// Mitsubishi GX Works2 project: 프로젝트1   PLC: Q03UDV

PROGRAM MAIN
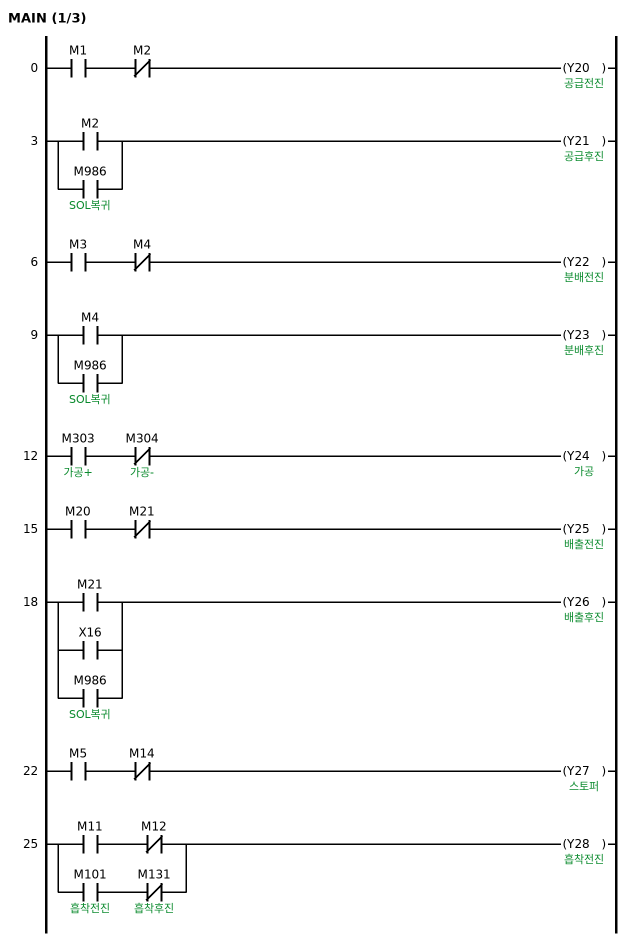
0     LD      M1
      ANI     M2
      OUT     Y20  ; 공급전진
3     LD      M2
      OR      M986  ; SOL복귀
      OUT     Y21  ; 공급후진
6     LD      M3
      ANI     M4
      OUT     Y22  ; 분배전진
9     LD      M4
      OR      M986  ; SOL복귀
      OUT     Y23  ; 분배후진
12    LD      M303  ; 가공+
      ANI     M304  ; 가공-
      OUT     Y24  ; 가공
15    LD      M20
      ANI     M21
      OUT     Y25  ; 배출전진
18    LD      M21
      OR      X16
      OR      M986  ; SOL복귀
      OUT     Y26  ; 배출후진
22    LD      M5
      ANI     M14
      OUT     Y27  ; 스토퍼
25    LD      M11
      ANI     M12
      LD      M101  ; 흡착전진
      ANI     M131  ; 흡착후진
      ORB
      OUT     Y28  ; 흡착전진
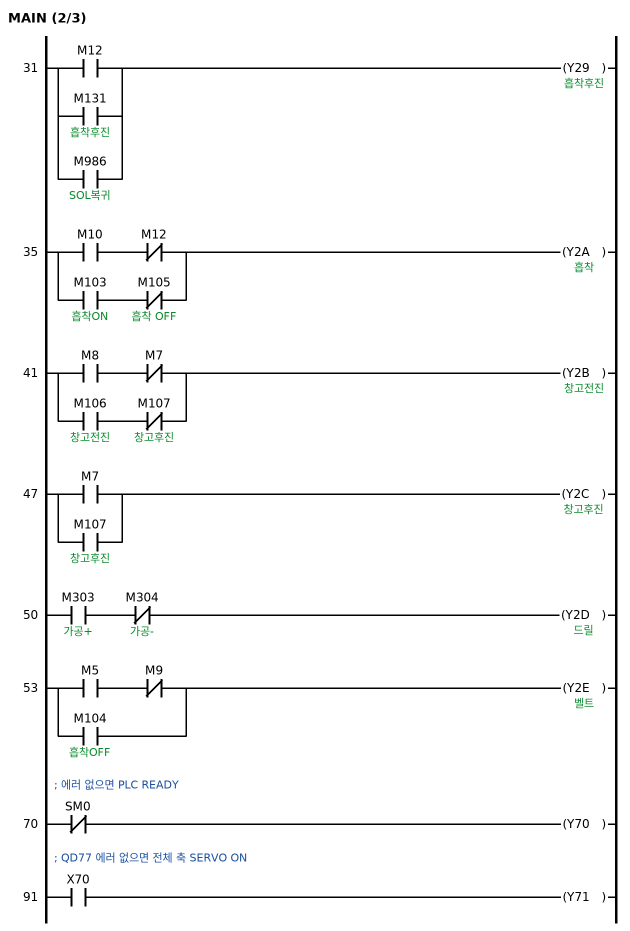
31    LD      M12
      OR      M131  ; 흡착후진
      OR      M986  ; SOL복귀
      OUT     Y29  ; 흡착후진
35    LD      M10
      ANI     M12
      LD      M103  ; 흡착ON
      ANI     M105  ; 흡착 OFF
      ORB
      OUT     Y2A  ; 흡착
41    LD      M8
      ANI     M7
      LD      M106  ; 창고전진
      ANI     M107  ; 창고후진
      ORB
      OUT     Y2B  ; 창고전진
47    LD      M7
      OR      M107  ; 창고후진
      OUT     Y2C  ; 창고후진
50    LD      M303  ; 가공+
      ANI     M304  ; 가공-
      OUT     Y2D  ; 드릴
53    LD      M5
      ANI     M9
      OR      M104  ; 흡착OFF
      OUT     Y2E  ; 벨트
; 에러 없으면 PLC READY
70    LDI     SM0
      OUT     Y70
; QD77 에러 없으면 전체 축 SERVO ON
91    LD      X70
      OUT     Y71
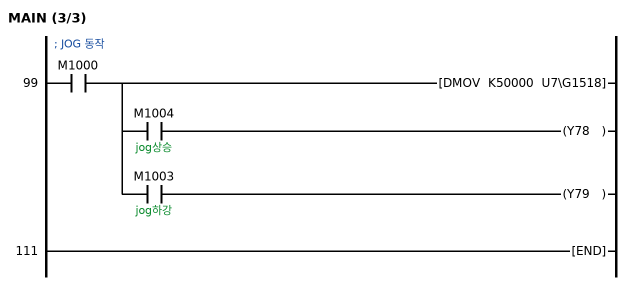
; JOG 동작
99    LD      M1000
      DMOV    K50000 U7\G1518
      MPS
      AND     M1004  ; jog상승
      OUT     Y78
      MPP
      AND     M1003  ; jog하강
      OUT     Y79
111   END
END_PROGRAM

PROGRAM OP
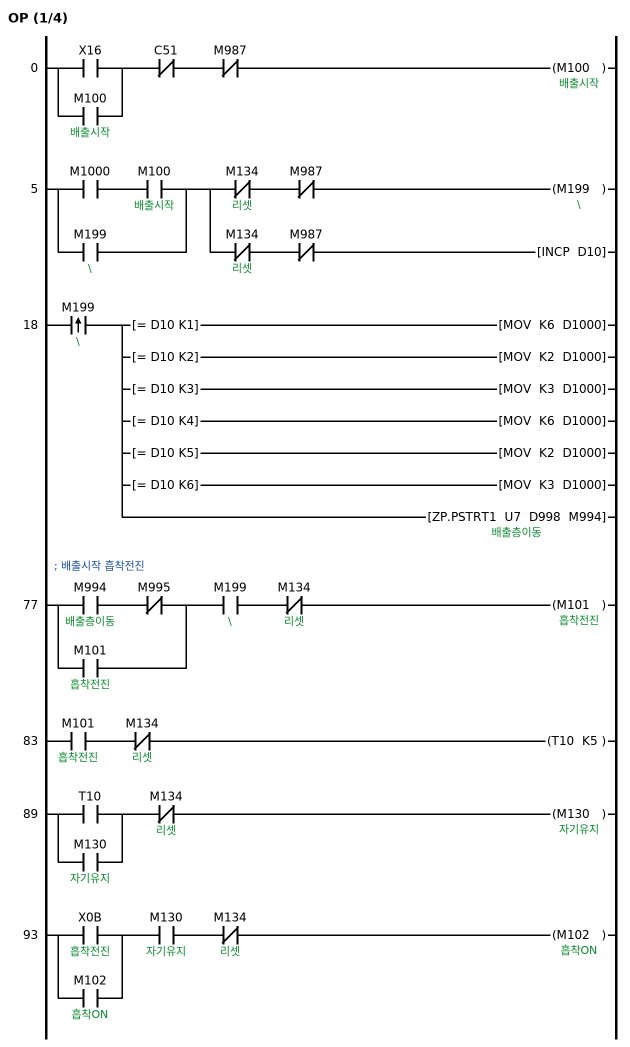
0     LD      X16
      OR      M100  ; 배출시작
      ANI     C51
      ANI     M987
      OUT     M100  ; 배출시작
5     LD      M1000
      AND     M100  ; 배출시작
      OR      M199  ; \
      MPS
      ANI     M134  ; 리셋
      ANI     M987
      OUT     M199  ; \
      MPP
      ANI     M134  ; 리셋
      ANI     M987
      INCP    D10
18    LDP     M199  ; \
      MPS
      AND=    D10 K1
      MOV     K6 D1000
      MRD
      AND=    D10 K2
      MOV     K2 D1000
      MRD
      AND=    D10 K3
      MOV     K3 D1000
      MRD
      AND=    D10 K4
      MOV     K6 D1000
      MRD
      AND=    D10 K5
      MOV     K2 D1000
      MRD
      AND=    D10 K6
      MOV     K3 D1000
      MPP
      ZP.PSTRT1 U7 D998 M994  ; 배출층이동
; 배출시작 흡착전진
77    LD      M994  ; 배출층이동
      ANI     M995
      OR      M101  ; 흡착전진
      AND     M199  ; \
      ANI     M134  ; 리셋
      OUT     M101  ; 흡착전진
83    LD      M101  ; 흡착전진
      ANI     M134  ; 리셋
      OUT     T10 K5
89    LD      T10
      OR      M130  ; 자기유지
      ANI     M134  ; 리셋
      OUT     M130  ; 자기유지
93    LD      X0B  ; 흡착전진
      OR      M102  ; 흡착ON
      AND     M130  ; 자기유지
      ANI     M134  ; 리셋
      OUT     M102  ; 흡착ON
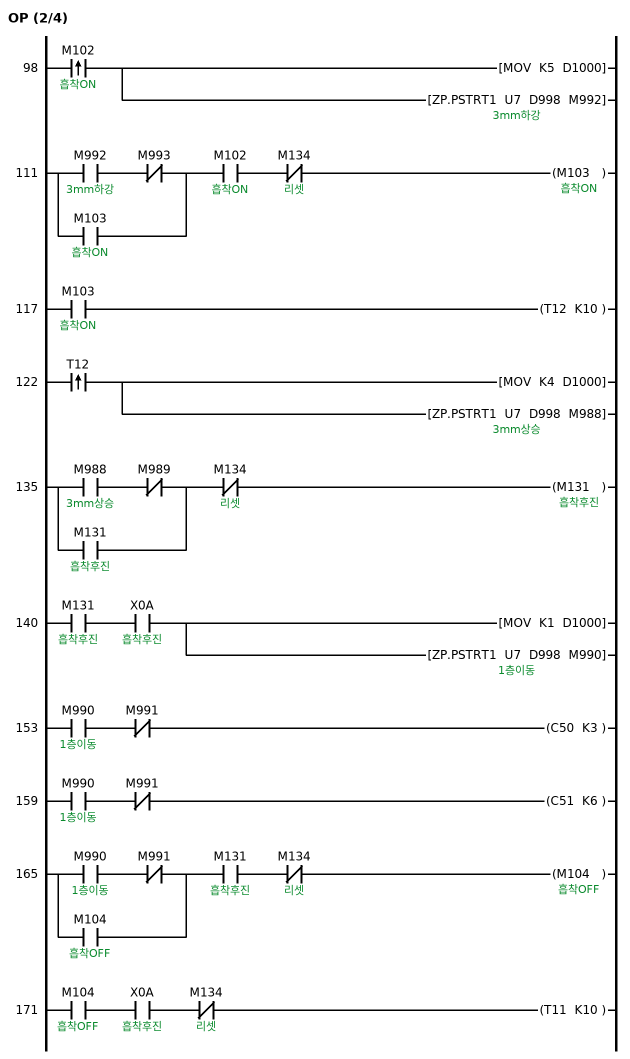
98    LDP     M102  ; 흡착ON
      MOV     K5 D1000
      ZP.PSTRT1 U7 D998 M992  ; 3mm하강
111   LD      M992  ; 3mm하강
      ANI     M993
      OR      M103  ; 흡착ON
      AND     M102  ; 흡착ON
      ANI     M134  ; 리셋
      OUT     M103  ; 흡착ON
117   LD      M103  ; 흡착ON
      OUT     T12 K10
122   LDP     T12
      MOV     K4 D1000
      ZP.PSTRT1 U7 D998 M988  ; 3mm상승
135   LD      M988  ; 3mm상승
      ANI     M989
      OR      M131  ; 흡착후진
      ANI     M134  ; 리셋
      OUT     M131  ; 흡착후진
140   LD      M131  ; 흡착후진
      AND     X0A  ; 흡착후진
      MOV     K1 D1000
      ZP.PSTRT1 U7 D998 M990  ; 1층이동
153   LD      M990  ; 1층이동
      ANI     M991
      OUT     C50 K3
159   LD      M990  ; 1층이동
      ANI     M991
      OUT     C51 K6
165   LD      M990  ; 1층이동
      ANI     M991
      OR      M104  ; 흡착OFF
      AND     M131  ; 흡착후진
      ANI     M134  ; 리셋
      OUT     M104  ; 흡착OFF
171   LD      M104  ; 흡착OFF
      AND     X0A  ; 흡착후진
      ANI     M134  ; 리셋
      OUT     T11 K10
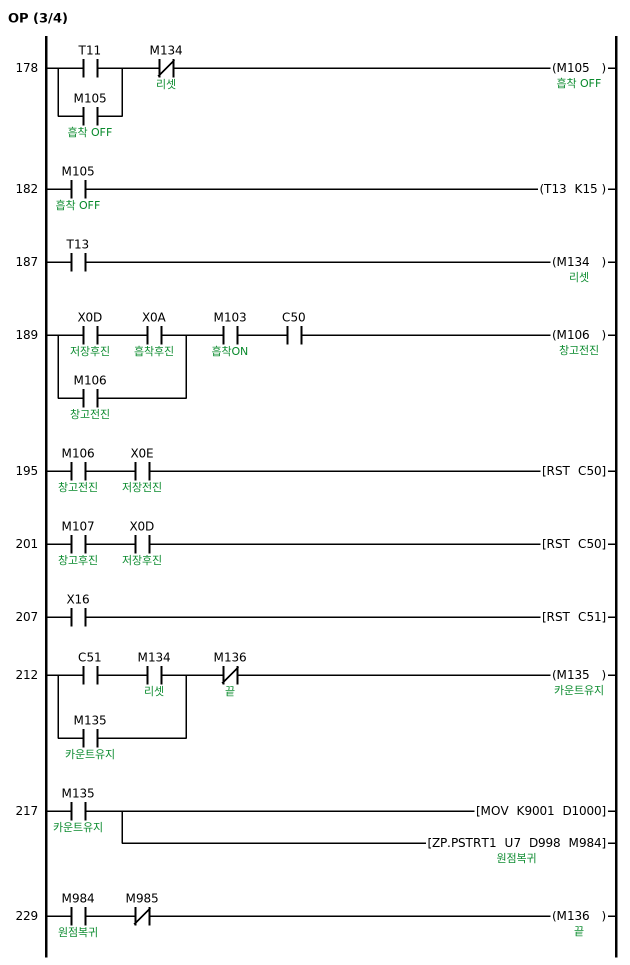
178   LD      T11
      OR      M105  ; 흡착 OFF
      ANI     M134  ; 리셋
      OUT     M105  ; 흡착 OFF
182   LD      M105  ; 흡착 OFF
      OUT     T13 K15
187   LD      T13
      OUT     M134  ; 리셋
189   LD      X0D  ; 저장후진
      AND     X0A  ; 흡착후진
      OR      M106  ; 창고전진
      AND     M103  ; 흡착ON
      AND     C50
      OUT     M106  ; 창고전진
195   LD      M106  ; 창고전진
      AND     X0E  ; 저장전진
      RST     C50
201   LD      M107  ; 창고후진
      AND     X0D  ; 저장후진
      RST     C50
207   LD      X16
      RST     C51
212   LD      C51
      AND     M134  ; 리셋
      OR      M135  ; 카운트유지
      ANI     M136  ; 끝
      OUT     M135  ; 카운트유지
217   LD      M135  ; 카운트유지
      MOV     K9001 D1000
      ZP.PSTRT1 U7 D998 M984  ; 원점복귀
229   LD      M984  ; 원점복귀
      ANI     M985
      OUT     M136  ; 끝
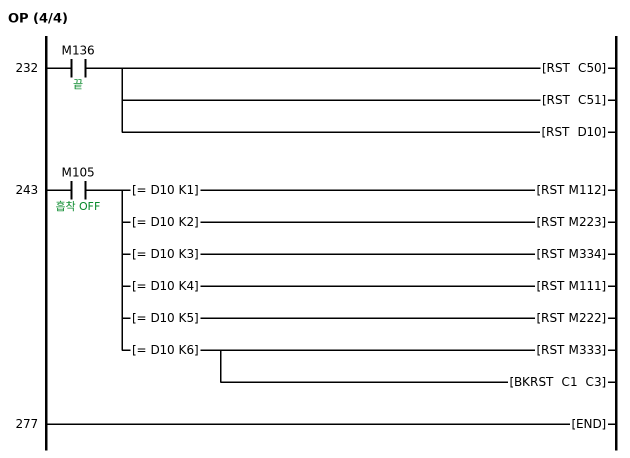
232   LD      M136  ; 끝
      RST     C50
      RST     C51
      RST     D10
243   LD      M105  ; 흡착 OFF
      MPS
      AND=    D10 K1
      RST     M112
      MRD
      AND=    D10 K2
      RST     M223
      MRD
      AND=    D10 K3
      RST     M334
      MRD
      AND=    D10 K4
      RST     M111
      MRD
      AND=    D10 K5
      RST     M222
      MPP
      AND=    D10 K6
      RST     M333
      BKRST   C1 C3
277   END
END_PROGRAM

PROGRAM MAIN1
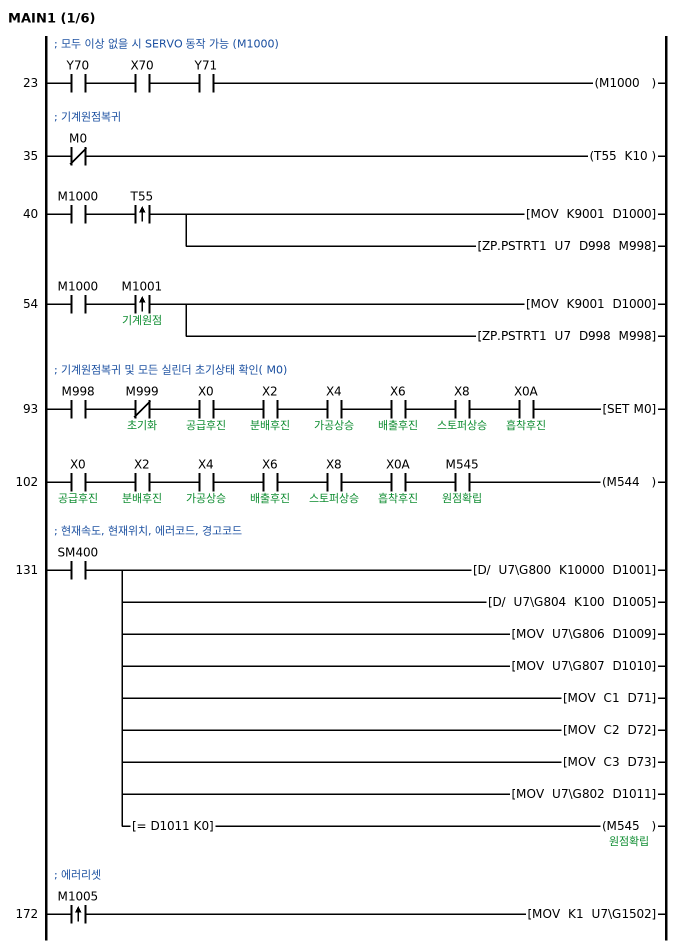
; 모두 이상 없을 시 SERVO 동작 가능 (M1000)
23    LD      Y70
      AND     X70
      AND     Y71
      OUT     M1000
; 기계원점복귀
35    LDI     M0
      OUT     T55 K10
40    LD      M1000
      ANDP    T55
      MOV     K9001 D1000
      ZP.PSTRT1 U7 D998 M998
54    LD      M1000
      ANDP    M1001  ; 기계원점
      MOV     K9001 D1000
      ZP.PSTRT1 U7 D998 M998
; 기계원점복귀 및 모든 실린더 초기상태 확인( M0)
93    LD      M998
      ANI     M999  ; 초기화
      AND     X0  ; 공급후진
      AND     X2  ; 분배후진
      AND     X4  ; 가공상승
      AND     X6  ; 배출후진
      AND     X8  ; 스토퍼상승
      AND     X0A  ; 흡착후진
      SET     M0
102   LD      X0  ; 공급후진
      AND     X2  ; 분배후진
      AND     X4  ; 가공상승
      AND     X6  ; 배출후진
      AND     X8  ; 스토퍼상승
      AND     X0A  ; 흡착후진
      AND     M545  ; 원점확립
      OUT     M544
; 현재속도, 현재위치, 에러코드, 경고코드
131   LD      SM400
      D/      U7\G800 K10000 D1001
      D/      U7\G804 K100 D1005
      MOV     U7\G806 D1009
      MOV     U7\G807 D1010
      MOV     C1 D71
      MOV     C2 D72
      MOV     C3 D73
      MOV     U7\G802 D1011
      AND=    D1011 K0
      OUT     M545  ; 원점확립
; 에러리셋
172   LDP     M1005
      MOV     K1 U7\G1502
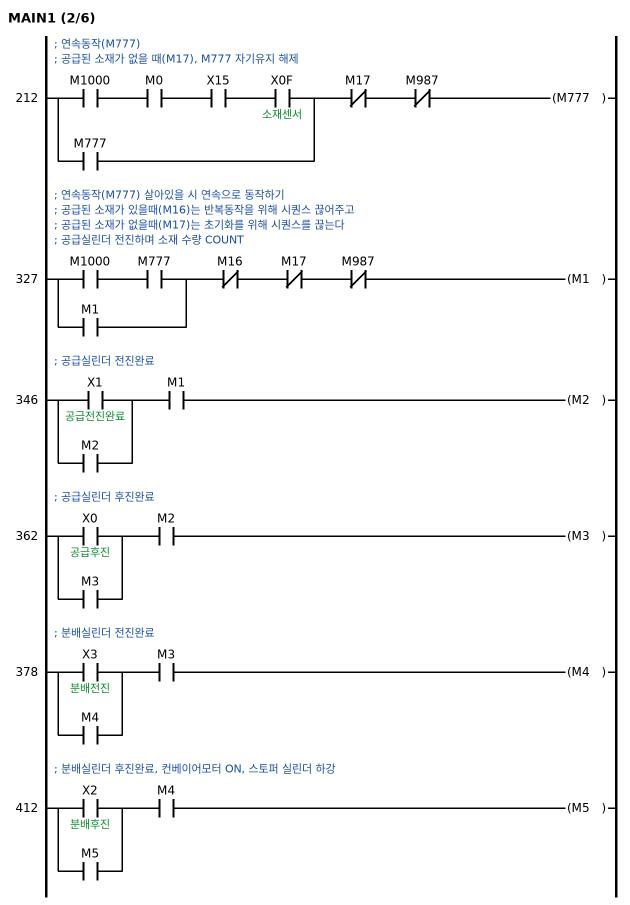
; 연속동작(M777)
; 공급된 소재가 없을 때(M17), M777 자기유지 해제
212   LD      M1000
      AND     M0
      AND     X15
      AND     X0F  ; 소재센서
      OR      M777
      ANI     M17
      ANI     M987
      OUT     M777
; 연속동작(M777) 살아있을 시 연속으로 동작하기
; 공급된 소재가 있을때(M16)는 반복동작을 위해 시퀀스 끊어주고
; 공급된 소재가 없을때(M17)는 초기화를 위해 시퀀스를 끊는다
; 공급실린더 전진하며 소재 수량 COUNT
327   LD      M1000
      AND     M777
      OR      M1
      ANI     M16
      ANI     M17
      ANI     M987
      OUT     M1
; 공급실린더 전진완료
346   LD      X1  ; 공급전진완료
      OR      M2
      AND     M1
      OUT     M2
; 공급실린더 후진완료
362   LD      X0  ; 공급후진
      OR      M3
      AND     M2
      OUT     M3
; 분배실린더 전진완료
378   LD      X3  ; 분배전진
      OR      M4
      AND     M3
      OUT     M4
; 분배실린더 후진완료, 컨베이어모터 ON, 스토퍼 실린더 하강
412   LD      X2  ; 분배후진
      OR      M5
      AND     M4
      OUT     M5
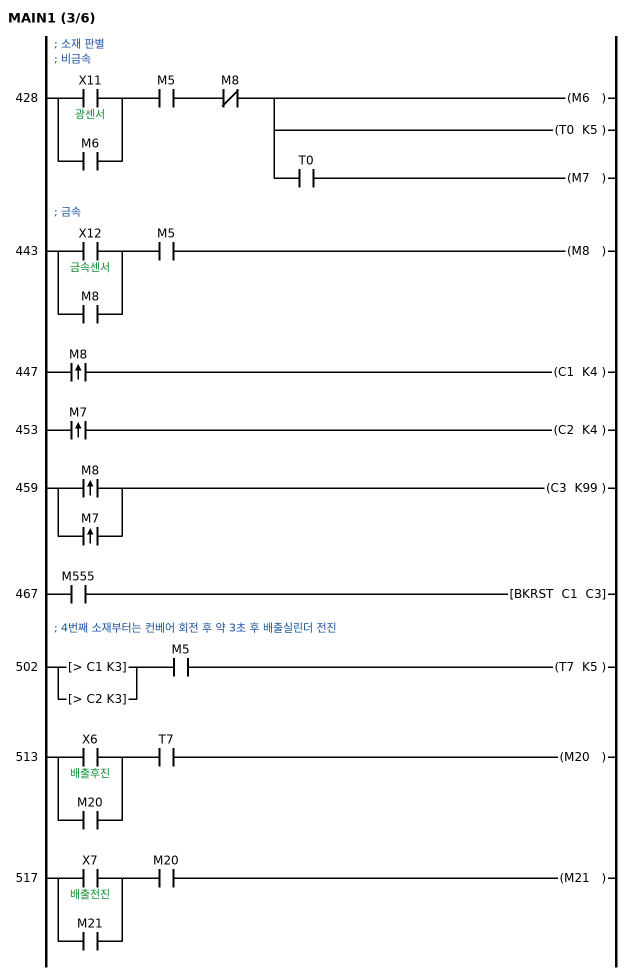
; 소재 판별
; 비금속
428   LD      X11  ; 광센서
      OR      M6
      AND     M5
      ANI     M8
      OUT     M6
      OUT     T0 K5
      AND     T0
      OUT     M7
; 금속
443   LD      X12  ; 금속센서
      OR      M8
      AND     M5
      OUT     M8
447   LDP     M8
      OUT     C1 K4
453   LDP     M7
      OUT     C2 K4
459   LDP     M8
      ORP     M7
      OUT     C3 K99
467   LD      M555
      BKRST   C1 C3
; 4번째 소재부터는 컨베어 회전 후 약 3초 후 배출실린더 전진
502   LD>     C1 K3
      OR>     C2 K3
      AND     M5
      OUT     T7 K5
513   LD      X6  ; 배출후진
      OR      M20
      AND     T7
      OUT     M20
517   LD      X7  ; 배출전진
      OR      M21
      AND     M20
      OUT     M21
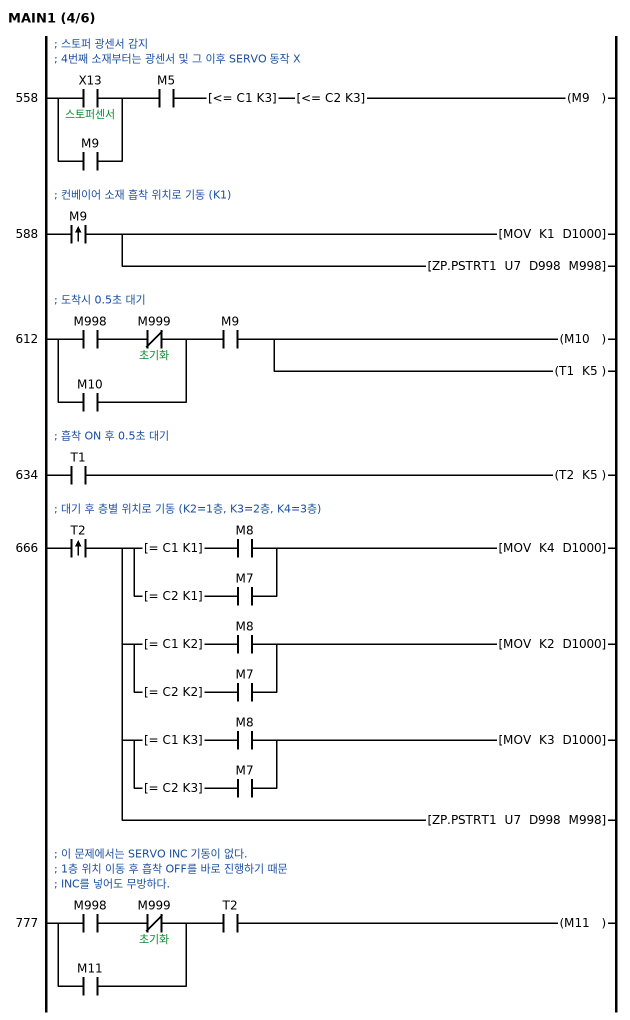
; 스토퍼 광센서 감지
; 4번째 소재부터는 광센서 및 그 이후 SERVO 동작 X
558   LD      X13  ; 스토퍼센서
      OR      M9
      AND     M5
      AND<=   C1 K3
      AND<=   C2 K3
      OUT     M9
; 컨베이어 소재 흡착 위치로 기동 (K1)
588   LDP     M9
      MOV     K1 D1000
      ZP.PSTRT1 U7 D998 M998
; 도착시 0.5초 대기
612   LD      M998
      ANI     M999  ; 초기화
      OR      M10
      AND     M9
      OUT     M10
      OUT     T1 K5
; 흡착 ON 후 0.5초 대기
634   LD      T1
      OUT     T2 K5
; 대기 후 층별 위치로 기동 (K2=1층, K3=2층, K4=3층)
666   LDP     T2
      MPS
      LD=     C1 K1
      AND     M8
      LD=     C2 K1
      AND     M7
      ORB
      ANB
      MOV     K4 D1000
      MRD
      LD=     C1 K2
      AND     M8
      LD=     C2 K2
      AND     M7
      ORB
      ANB
      MOV     K2 D1000
      MRD
      LD=     C1 K3
      AND     M8
      LD=     C2 K3
      AND     M7
      ORB
      ANB
      MOV     K3 D1000
      MPP
      ZP.PSTRT1 U7 D998 M998
; 이 문제에서는 SERVO INC 기동이 없다.
; 1층 위치 이동 후 흡착 OFF를 바로 진행하기 때문
; INC를 넣어도 무방하다.
777   LD      M998
      ANI     M999  ; 초기화
      OR      M11
      AND     T2
      OUT     M11
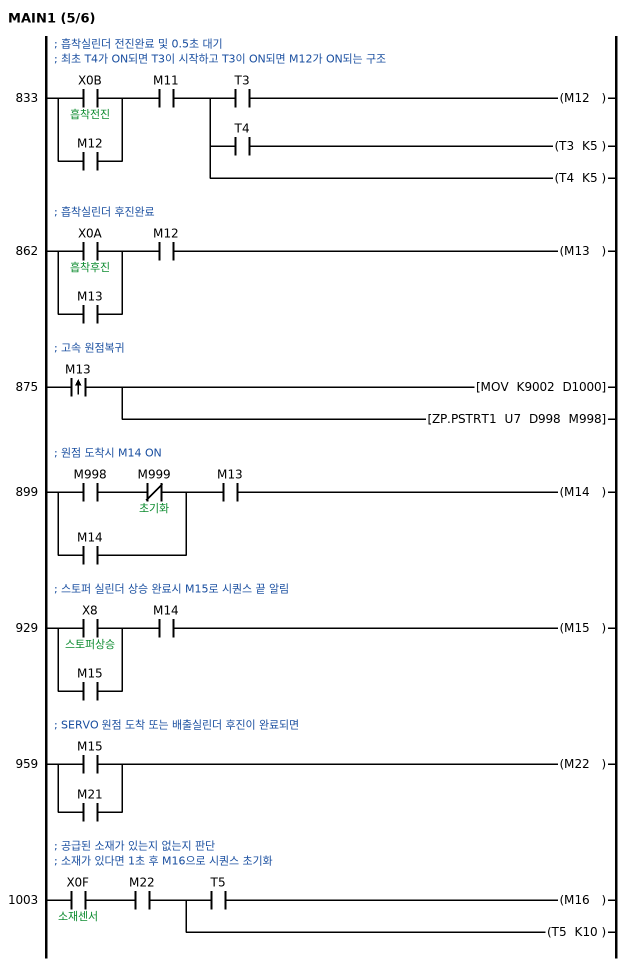
; 흡착실린더 전진완료 및 0.5초 대기
; 최초 T4가 ON되면 T3이 시작하고 T3이 ON되면 M12가 ON되는 구조
833   LD      X0B  ; 흡착전진
      OR      M12
      AND     M11
      MPS
      AND     T3
      OUT     M12
      MRD
      AND     T4
      OUT     T3 K5
      MPP
      OUT     T4 K5
; 흡착실린더 후진완료
862   LD      X0A  ; 흡착후진
      OR      M13
      AND     M12
      OUT     M13
; 고속 원점복귀
875   LDP     M13
      MOV     K9002 D1000
      ZP.PSTRT1 U7 D998 M998
; 원점 도착시 M14 ON
899   LD      M998
      ANI     M999  ; 초기화
      OR      M14
      AND     M13
      OUT     M14
; 스토퍼 실린더 상승 완료시 M15로 시퀀스 끝 알림
929   LD      X8  ; 스토퍼상승
      OR      M15
      AND     M14
      OUT     M15
; SERVO 원점 도착 또는 배출실린더 후진이 완료되면
959   LD      M15
      OR      M21
      OUT     M22
; 공급된 소재가 있는지 없는지 판단
; 소재가 있다면 1초 후 M16으로 시퀀스 초기화
1003  LD      X0F  ; 소재센서
      AND     M22
      MPS
      AND     T5
      OUT     M16
      MPP
      OUT     T5 K10
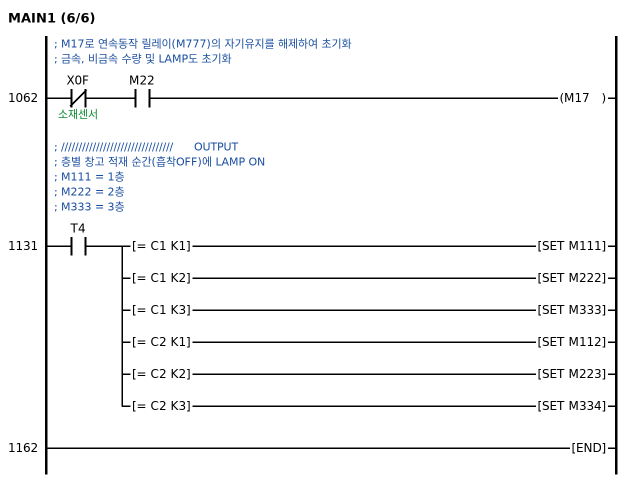
; M17로 연속동작 릴레이(M777)의 자기유지를 해제하여 초기화
; 금속, 비금속 수량 및 LAMP도 초기화
1062  LDI     X0F  ; 소재센서
      AND     M22
      OUT     M17
; ////////////////////////////////      OUTPUT
; 층별 창고 적재 순간(흡착OFF)에 LAMP ON
; M111 = 1층
; M222 = 2층
; M333 = 3층
1131  LD      T4
      MPS
      AND=    C1 K1
      SET     M111
      MRD
      AND=    C1 K2
      SET     M222
      MRD
      AND=    C1 K3
      SET     M333
      MRD
      AND=    C2 K1
      SET     M112
      MRD
      AND=    C2 K2
      SET     M223
      MPP
      AND=    C2 K3
      SET     M334
1162  END
END_PROGRAM

// device comments not shown above
X5  ; 가공하강
M50  ; 정상속도
M51  ; 비정상속도
M300  ; 작동
M301  ; 공급+
M302  ; 공급-
M305  ; 카운트
M306  ; 가공카운트
M307  ; 분배+
M308  ; 분배-
M309  ; 벨트+
M310  ; 스토퍼+
M311  ; 벨트정지
M312  ; 1층후흡착
M313  ; 흡착후up
M314  ; 흡착전진
M315  ; 1층적재
M316  ; 흡착후진
M318  ; 1층완료
M319  ; 2층전진
M320  ; 2층흡착/
M321  ; 2층후진
M323  ; 저장후진ㄱ
M324  ; 저장전진
M325  ; 2층완료
M326  ; 벨트흡착2
M327  ; 흡착후UP
M328  ; 소재판단
M329  ; 스토퍼유지
M330  ; 스토퍼유지
M331  ; 흡착전진2
M332  ; 흡착후진
M336  ; 흡착ON
M395  ; 카운트완
M396  ; 카운트
M397  ; 가공-
M398  ; 가공+
M400  ; 1층도착
M402  ; 3mmUP
M404  ; 원점복귀
M406  ; 2층보냄
M408  ; 2층적재후복귀
M410  ; 2층후복귀
M888  ; reset
M1002  ; 고속원점
T6  ; 0.5초
C13  ; 2회
